{attribute 'qualified_only'}
{attribute 'strict'}
{attribute 'to_string'}
TYPE E_Led_Color :
(
	Yellow := 0,
	Red,
	Green,
	Blue,
	Gray
	
);
END_TYPE

(* stored: Version 1.1.0.1, ProductVersion 3.1.4024.12
   DUT E_Led_Color: Id {8e307ad3-6cdf-4023-85ee-14ef20693336} *)
